(* PLC project Claude2.project, CODESYS CODESYS V3.5 SP20 *)
(* stored: creationDateTime 2026-10-26T14:12:36.8389124, modificationDateTime 2026-10-26T14:11:59.3278775 *)

(* values of E_MachineState: INIT: Inicialização; STOPPED: Parada, sem alarme; HOMING: Referenciamento dos eixos; RUNNING: Ciclo automático; ALARM: Alarme pendente: parada segura; ESTOP: Emergência/porta aberta: sobrepõe tudo *)

{attribute 'qualified_only'}
{attribute 'strict'}
TYPE E_MachineState : (INIT := 0, STOPPED := 10, HOMING := 20, RUNNING := 30, ALARM := 90, ESTOP := 99);
END_TYPE

TYPE ST_Component : STRUCT
  sRef : STRING(20);  (* Designador do componente *)
  rPickX : REAL;  (* Posição de coleta (alimentador) X [mm] *)
  rPickY : REAL;  (* Posição de coleta (alimentador) Y [mm] *)
  rPlaceX : REAL;  (* Posição de montagem X [mm] *)
  rPlaceY : REAL;  (* Posição de montagem Y [mm] *)
  rPlaceTheta : REAL;  (* Ângulo de montagem [graus] *)
END_STRUCT;
END_TYPE

TYPE ST_Recipe : STRUCT
  sName : STRING(30);  (* Nome da receita *)
  iCount : INT;  (* Quantidade de componentes *)
  aComp : ARRAY[1..c_MAX_COMP] OF ST_Component;  (* Lista de componentes *)
END_STRUCT;
END_TYPE

FUNCTION F_InRange : BOOL
  VAR_INPUT
    rValue : REAL;
    rMin : REAL;
    rMax : REAL;
  END_VAR

                  (* Verifica se o valor está dentro da faixa [rMin, rMax] *)
F_InRange := (rValue >= rMin) AND (rValue <= rMax);
                
END_FUNCTION

FUNCTION_BLOCK FB_PneumaticCyl
  VAR_INPUT
    xEnable : BOOL;  (* Habilitação (segurança) *)
    xReset : BOOL;  (* Reset de falha *)
    xCmdExtend : BOOL;  (* TRUE = avançar; FALSE = recuar *)
    xSensExtended : BOOL;
    xSensRetracted : BOOL;
    tMoveTimeout : TIME := TIME#2s0ms;
    tSensorConflict : TIME := TIME#300ms;
  END_VAR
  VAR_OUTPUT
    xValve : BOOL;
    xIsExtended : BOOL;  (* Avançado confirmado: sensor A ligado e B desligado *)
    xIsRetracted : BOOL;  (* Recuado confirmado: sensor B ligado e A desligado *)
    xFault : BOOL;
    iFaultCode : INT;  (* 1 = timeout avanço; 2 = timeout recuo; 3 = sensores em conflito *)
  END_VAR
  VAR
    tonExt : TON;
    tonRet : TON;
    tonBoth : TON;
  END_VAR

                  (* Dupla confirmação *)
xIsExtended  := xSensExtended AND NOT xSensRetracted;
xIsRetracted := xSensRetracted AND NOT xSensExtended;

IF xReset THEN
    xFault := FALSE;
    iFaultCode := 0;
END_IF

(* Supervisão de tempo e de coerência dos sensores *)
tonExt(IN := xEnable AND xValve AND NOT xIsExtended AND NOT xFault, PT := tMoveTimeout);
tonRet(IN := xEnable AND NOT xValve AND NOT xIsRetracted AND NOT xFault, PT := tMoveTimeout);
tonBoth(IN := xEnable AND xSensExtended AND xSensRetracted, PT := tSensorConflict);

IF NOT xFault THEN
    IF tonExt.Q THEN
        xFault := TRUE; iFaultCode := 1;
    ELSIF tonRet.Q THEN
        xFault := TRUE; iFaultCode := 2;
    ELSIF tonBoth.Q THEN
        xFault := TRUE; iFaultCode := 3;
    END_IF
END_IF

(* Saída da válvula: em falha ou sem habilitação, retorna por mola *)
xValve := xEnable AND xCmdExtend AND NOT xFault;
                
END_FUNCTION_BLOCK

FUNCTION_BLOCK FB_VacuumGripper
  VAR_INPUT
    xEnable : BOOL;
    xReset : BOOL;
    xGrip : BOOL;  (* TRUE = segurar; FALSE = liberar *)
    xPressostat : BOOL;
    tConfirm : TIME := TIME#1s0ms;  (* Tempo máximo para confirmar a pega *)
    tDebounce : TIME := TIME#100ms;
    tBlow : TIME := TIME#300ms;
  END_VAR
  VAR_OUTPUT
    xVacValve : BOOL;
    xBlowValve : BOOL;
    xGripOk : BOOL;  (* Pega confirmada *)
    xReleased : BOOL;  (* Liberação confirmada *)
    xPickFail : BOOL;  (* Pega não confirmada no tempo *)
    xGripLoss : BOOL;  (* Perda de vácuo com peça presa *)
  END_VAR
  VAR
    tonOk : TON;
    tonConfirm : TON;
    tonLoss : TON;
    tonRel : TON;
    tonBlow : TON;
    ftGrip : F_TRIG;
    xBlow : BOOL;
    xCarried : BOOL;
  END_VAR

                  xVacValve := xEnable AND xGrip;

(* Janela de sopro após o comando de liberação *)
ftGrip(CLK := xGrip);
IF ftGrip.Q THEN
    xBlow := TRUE;
END_IF
tonBlow(IN := xBlow, PT := tBlow);
IF tonBlow.Q OR xGrip OR NOT xEnable THEN
    xBlow := FALSE;
END_IF
xBlowValve := xBlow AND xEnable;

(* Confirmação da pega *)
tonOk(IN := xGrip AND xPressostat, PT := tDebounce);
xGripOk := tonOk.Q;

(* Falha de pega: vácuo não estabelecido no tempo *)
tonConfirm(IN := xEnable AND xGrip AND NOT xGripOk, PT := tConfirm);
IF tonConfirm.Q THEN
    xPickFail := TRUE;
END_IF
IF xReset OR NOT xGrip THEN
    xPickFail := FALSE;
END_IF

(* Perda de vácuo durante o transporte *)
IF xGripOk THEN
    xCarried := TRUE;
END_IF
IF NOT xGrip THEN
    xCarried := FALSE;
END_IF
tonLoss(IN := xCarried AND xGrip AND NOT xPressostat, PT := tDebounce);
xGripLoss := tonLoss.Q;

(* Confirmação da liberação *)
tonRel(IN := NOT xGrip AND NOT xPressostat, PT := tDebounce);
xReleased := tonRel.Q;
                
END_FUNCTION_BLOCK

FUNCTION_BLOCK FB_AxisCtrl
  VAR_INPUT
    xEnable : BOOL;
    xReset : BOOL;
    xHomeCmd : BOOL;  (* Borda de subida inicia o homing *)
    xMoveCmd : BOOL;  (* Borda de subida inicia o movimento *)
    xHalt : BOOL;  (* Interrompe o movimento em curso *)
    rTarget : REAL;
    rActPos : REAL;
    rSoftMin : REAL;
    rSoftMax : REAL;
    xDriveReady : BOOL;
    xDriveFault : BOOL;
    xDriveHomeDone : BOOL;
    rInPosWindow : REAL := 0.05;
    tSettle : TIME := TIME#100ms;
    tReadyTimeout : TIME := TIME#5s0ms;
    tHomeTimeout : TIME := TIME#1m0s0ms;
    tMoveTimeout : TIME := TIME#15s0ms;
  END_VAR
  VAR_OUTPUT
    xDrivePower : BOOL;
    xDriveHome : BOOL;
    xDriveExecute : BOOL;  (* Pulso de um ciclo *)
    rDriveSetpoint : REAL;
    xHomed : BOOL;
    xInPos : BOOL;
    xBusy : BOOL;
    xAccept : BOOL;  (* Apto a receber comando de homing/movimento *)
    xFault : BOOL;
    iFaultCode : INT;  (* 1 drive não pronto; 2 timeout homing; 3 alvo fora dos limites; 4 timeout movimento; 5 falha do drive; 6 perda de pronto *)
  END_VAR
  VAR
    iState : INT := 0;
    rtHome : R_TRIG;
    rtMove : R_TRIG;
    tonReady : TON;
    tonHome : TON;
    tonMove : TON;
    tonSettle : TON;
    rLastSetpoint : REAL;
    rLatchTarget : REAL;
    xHaltDone : BOOL;
  END_VAR
  VAR CONSTANT
    AS_OFF : INT := 0;
    AS_WAIT_READY : INT := 1;
    AS_UNHOMED : INT := 2;
    AS_HOMING : INT := 3;
    AS_READY : INT := 4;
    AS_START : INT := 5;
    AS_MOVING : INT := 6;
    AS_FAULT : INT := 99;
  END_VAR

                  xDriveExecute := FALSE;
rtHome(CLK := xHomeCmd);
rtMove(CLK := xMoveCmd);

tonReady(IN := (iState = AS_WAIT_READY), PT := tReadyTimeout);
tonHome(IN := (iState = AS_HOMING), PT := tHomeTimeout);
tonMove(IN := (iState = AS_MOVING), PT := tMoveTimeout);
tonSettle(IN := (iState = AS_MOVING) AND (ABS(rActPos - rLastSetpoint) <= rInPosWindow),
          PT := tSettle);

(* Supervisão geral *)
IF iState <> AS_FAULT THEN
    IF NOT xEnable THEN
        iState := AS_OFF;
    ELSIF iState >= AS_WAIT_READY THEN
        IF xDriveFault THEN
            iFaultCode := 5; iState := AS_FAULT;
        ELSIF (iState >= AS_UNHOMED) AND NOT xDriveReady THEN
            iFaultCode := 6; iState := AS_FAULT;
        END_IF
    END_IF
END_IF

CASE iState OF
    AS_OFF:
        xHomed := FALSE;
        IF xEnable THEN
            iState := AS_WAIT_READY;
        END_IF

    AS_WAIT_READY:
        IF xDriveReady THEN
            iState := AS_UNHOMED;
        ELSIF tonReady.Q THEN
            iFaultCode := 1; iState := AS_FAULT;
        END_IF

    AS_UNHOMED:
        IF rtHome.Q THEN
            iState := AS_HOMING;
        END_IF

    AS_HOMING:
        IF xDriveHomeDone THEN
            xHomed := TRUE;
            rLastSetpoint := rActPos;
            iState := AS_READY;
        ELSIF tonHome.Q THEN
            iFaultCode := 2; iState := AS_FAULT;
        END_IF

    AS_READY:
        IF rtHome.Q THEN
            xHomed := FALSE;
            iState := AS_HOMING;
        ELSIF rtMove.Q THEN
            IF (rTarget < rSoftMin) OR (rTarget > rSoftMax) THEN
                iFaultCode := 3; iState := AS_FAULT;
            ELSE
                rLatchTarget := rTarget;
                iState := AS_START;
            END_IF
        END_IF

    AS_START:
        rDriveSetpoint := rLatchTarget;
        rLastSetpoint := rLatchTarget;
        xDriveExecute := TRUE;
        iState := AS_MOVING;

    AS_MOVING:
        IF xHalt AND NOT xHaltDone THEN
            (* Parada: novo alvo = posição atual *)
            rDriveSetpoint := rActPos;
            rLastSetpoint := rActPos;
            xDriveExecute := TRUE;
            xHaltDone := TRUE;
        END_IF
        IF tonSettle.Q THEN
            iState := AS_READY;
        ELSIF tonMove.Q THEN
            iFaultCode := 4; iState := AS_FAULT;
        END_IF

    AS_FAULT:
        xHomed := FALSE;
        IF xReset AND NOT xDriveFault THEN
            iFaultCode := 0;
            iState := AS_OFF;
        END_IF
END_CASE

IF iState <> AS_MOVING THEN
    xHaltDone := FALSE;
END_IF

(* Saídas *)
xDrivePower := (iState >= AS_WAIT_READY) AND (iState <> AS_FAULT);
xDriveHome  := (iState = AS_HOMING);
xBusy       := (iState = AS_HOMING) OR (iState = AS_START) OR (iState = AS_MOVING);
xAccept     := (iState = AS_UNHOMED) OR (iState = AS_READY);
xInPos      := (iState = AS_READY) AND xHomed AND (ABS(rActPos - rLastSetpoint) <= rInPosWindow);
xFault      := (iState = AS_FAULT);
                
END_FUNCTION_BLOCK

FUNCTION_BLOCK FB_Conveyor
  VAR_INPUT
    xEnable : BOOL;  (* Ciclo automático liberado *)
    xReset : BOOL;
    xClearZones : BOOL;  (* Ressincroniza zonas pelos sensores *)
    xSensZ1 : BOOL;
    xSensZ2 : BOOL;
    xSensZ3 : BOOL;
    xUpBoardAvail : BOOL;  (* SMEMA a montante: placa disponível *)
    xDownMachineReady : BOOL;  (* SMEMA a jusante: máquina pronta *)
    xAsmDone : BOOL;  (* Montagem concluída: libera a zona 2 *)
    xInspDone : BOOL;  (* Inspeção concluída: libera a zona 3 *)
    tTransferTimeout : TIME := TIME#15s0ms;
    tSensorFilter : TIME := TIME#50ms;
    tClearDelay : TIME := TIME#500ms;
  END_VAR
  VAR_OUTPUT
    xMotor1 : BOOL;
    xMotor2 : BOOL;
    xMotor3 : BOOL;
    xUpMachineReady : BOOL;  (* SMEMA a montante: máquina pronta *)
    xDownBoardAvail : BOOL;  (* SMEMA a jusante: placa disponível *)
    xBoardInAsm : BOOL;
    xBoardInInsp : BOOL;
    xFault : BOOL;
  END_VAR
  VAR
    iZ1 : INT;  (* Estado de cada zona *)
    iZ2 : INT;  (* Estado de cada zona *)
    iZ3 : INT;  (* Estado de cada zona *)
    tonP1 : TON;  (* Presença filtrada *)
    tonP2 : TON;  (* Presença filtrada *)
    tonP3 : TON;  (* Presença filtrada *)
    tonA1 : TON;  (* Ausência filtrada *)
    tonA2 : TON;  (* Ausência filtrada *)
    tonA3 : TON;  (* Ausência filtrada *)
    tonT1 : TON;  (* Timeout de movimento *)
    tonT2 : TON;  (* Timeout de movimento *)
    tonT3 : TON;  (* Timeout de movimento *)
    xP1 : BOOL;
    xP2 : BOOL;
    xP3 : BOOL;
    xA1 : BOOL;
    xA2 : BOOL;
    xA3 : BOOL;
    xActive : BOOL;
  END_VAR
  VAR CONSTANT
    ZS_EMPTY : INT := 0;
    ZS_RECV : INT := 1;  (* Recebendo placa *)
    ZS_OCC : INT := 2;  (* Placa posicionada *)
    ZS_SEND : INT := 3;  (* Enviando placa *)
  END_VAR

                  (* Filtros dos sensores *)
tonP1(IN := xSensZ1, PT := tSensorFilter);   xP1 := tonP1.Q;
tonP2(IN := xSensZ2, PT := tSensorFilter);   xP2 := tonP2.Q;
tonP3(IN := xSensZ3, PT := tSensorFilter);   xP3 := tonP3.Q;
tonA1(IN := NOT xSensZ1, PT := tClearDelay); xA1 := tonA1.Q;
tonA2(IN := NOT xSensZ2, PT := tClearDelay); xA2 := tonA2.Q;
tonA3(IN := NOT xSensZ3, PT := tClearDelay); xA3 := tonA3.Q;

IF xReset THEN
    xFault := FALSE;
END_IF

(* Ressincronização: considera placa posicionada onde houver sensor ativo *)
IF xClearZones THEN
    IF xSensZ1 THEN iZ1 := ZS_OCC; ELSE iZ1 := ZS_EMPTY; END_IF
    IF xSensZ2 THEN iZ2 := ZS_OCC; ELSE iZ2 := ZS_EMPTY; END_IF
    IF xSensZ3 THEN iZ3 := ZS_OCC; ELSE iZ3 := ZS_EMPTY; END_IF
    xFault := FALSE;
END_IF

(* Timeout de transferência (motores acionados no ciclo anterior) *)
tonT1(IN := xMotor1, PT := tTransferTimeout);
tonT2(IN := xMotor2, PT := tTransferTimeout);
tonT3(IN := xMotor3, PT := tTransferTimeout);
IF tonT1.Q OR tonT2.Q OR tonT3.Q THEN
    xFault := TRUE;
END_IF

xActive := xEnable AND NOT xFault;

(* ---------- Zona 1: entrada ---------- *)
CASE iZ1 OF
    ZS_EMPTY:
        IF xActive AND xUpBoardAvail THEN
            iZ1 := ZS_RECV;
        END_IF
    ZS_RECV:
        IF xP1 THEN
            iZ1 := ZS_OCC;
        END_IF
    ZS_OCC:
        IF xActive AND (iZ2 = ZS_EMPTY) THEN
            iZ1 := ZS_SEND;
            iZ2 := ZS_RECV;     (* Transferência 1 -> 2 *)
        END_IF
    ZS_SEND:
        IF (iZ2 = ZS_OCC) AND xA1 THEN
            iZ1 := ZS_EMPTY;
        END_IF
END_CASE

(* ---------- Zona 2: montagem ---------- *)
CASE iZ2 OF
    ZS_EMPTY:
        ;
    ZS_RECV:
        IF xP2 THEN
            iZ2 := ZS_OCC;
        END_IF
    ZS_OCC:
        IF xActive AND xAsmDone AND (iZ3 = ZS_EMPTY) THEN
            iZ2 := ZS_SEND;
            iZ3 := ZS_RECV;     (* Transferência 2 -> 3 *)
        END_IF
    ZS_SEND:
        IF (iZ3 = ZS_OCC) AND xA2 THEN
            iZ2 := ZS_EMPTY;
        END_IF
END_CASE

(* ---------- Zona 3: saída / inspeção ---------- *)
CASE iZ3 OF
    ZS_EMPTY:
        ;
    ZS_RECV:
        IF xP3 THEN
            iZ3 := ZS_OCC;
        END_IF
    ZS_OCC:
        IF xActive AND xInspDone THEN
            iZ3 := ZS_SEND;
        END_IF
    ZS_SEND:
        IF xA3 THEN
            iZ3 := ZS_EMPTY;
        END_IF
END_CASE

(* ---------- Saídas (calculadas após a lógica de estados) ---------- *)
xMotor1 := xActive AND ((iZ1 = ZS_RECV) OR (iZ1 = ZS_SEND));
xMotor2 := xActive AND ((iZ2 = ZS_RECV) OR (iZ2 = ZS_SEND));
xMotor3 := xActive AND ((iZ3 = ZS_RECV) OR ((iZ3 = ZS_SEND) AND xDownMachineReady));

xUpMachineReady := xActive AND ((iZ1 = ZS_EMPTY) OR (iZ1 = ZS_RECV));
xDownBoardAvail := (iZ3 = ZS_SEND);
xBoardInAsm     := (iZ2 = ZS_OCC);
xBoardInInsp    := (iZ3 = ZS_OCC);
                
END_FUNCTION_BLOCK

FUNCTION_BLOCK FB_HmiWatchdog
  VAR_INPUT
    iHeartbeat : UINT;
    tTimeout : TIME := TIME#3s0ms;
  END_VAR
  VAR_OUTPUT
    xOk : BOOL;
    xLost : BOOL;
  END_VAR
  VAR
    uiLast : UINT;
    xFirst : BOOL := TRUE;
    xChanged : BOOL;
    tonLoss : TON;
  END_VAR

                  IF xFirst THEN
    uiLast := iHeartbeat;
    xFirst := FALSE;
END_IF

xChanged := (iHeartbeat <> uiLast);
uiLast := iHeartbeat;

tonLoss(IN := NOT xChanged, PT := tTimeout);
xLost := tonLoss.Q;
xOk := NOT tonLoss.Q;
                
END_FUNCTION_BLOCK

FUNCTION_BLOCK FB_Alarm
  VAR_INPUT
    xCondition : BOOL;  (* Condição de alarme (nível ou pulso) *)
    xAck : BOOL;
    xReset : BOOL;
  END_VAR
  VAR_OUTPUT
    xActive : BOOL;  (* Alarme retido *)
    xAcked : BOOL;
  END_VAR
  VAR
    rtCond : R_TRIG;
    rtAck : R_TRIG;
    rtRst : R_TRIG;
  END_VAR

                  rtCond(CLK := xCondition);
rtAck(CLK := xAck);
rtRst(CLK := xReset);

IF rtCond.Q THEN
    xActive := TRUE;
    xAcked := FALSE;
END_IF

IF rtAck.Q AND xActive THEN
    xAcked := TRUE;
END_IF

(* Reset só é aceito com alarme reconhecido e condição normalizada *)
IF rtRst.Q AND xActive AND xAcked AND NOT xCondition THEN
    xActive := FALSE;
    xAcked := FALSE;
END_IF
                
END_FUNCTION_BLOCK

FUNCTION_BLOCK FB_Recipe
  VAR_INPUT
    xRequest : BOOL;  (* Borda de subida solicita a troca *)
    iRequested : INT;
    xMachineStopped : BOOL;
    rXMin : REAL;
    rXMax : REAL;
    rYMin : REAL;
    rYMax : REAL;
  END_VAR
  VAR_IN_OUT
    aRecipes : ARRAY[1..c_NUM_RECIPES] OF ST_Recipe;
  END_VAR
  VAR_OUTPUT
    iActive : INT;
    xValid : BOOL;
    xRejected : BOOL;
  END_VAR
  VAR
    rtReq : R_TRIG;
    i : INT;
    xOk : BOOL;
    stC : ST_Component;
  END_VAR

                  rtReq(CLK := xRequest);

IF rtReq.Q THEN
    IF xMachineStopped AND (iRequested >= 1) AND (iRequested <= c_NUM_RECIPES) THEN
        iActive := iRequested;
        xRejected := FALSE;
    ELSE
        xRejected := TRUE;
    END_IF
END_IF
IF NOT xRequest THEN
    xRejected := FALSE;
END_IF

(* Validação da receita ativa *)
xOk := (iActive >= 1) AND (iActive <= c_NUM_RECIPES);
IF xOk THEN
    xOk := (aRecipes[iActive].iCount >= 1) AND (aRecipes[iActive].iCount <= c_MAX_COMP);
END_IF
IF xOk THEN
    FOR i := 1 TO aRecipes[iActive].iCount DO
        stC := aRecipes[iActive].aComp[i];
        IF NOT (F_InRange(stC.rPickX, rXMin, rXMax)
            AND F_InRange(stC.rPickY, rYMin, rYMax)
            AND F_InRange(stC.rPlaceX, rXMin, rXMax)
            AND F_InRange(stC.rPlaceY, rYMin, rYMax)
            AND F_InRange(stC.rPlaceTheta, -180.0, 180.0)) THEN
            xOk := FALSE;
            EXIT;
        END_IF
    END_FOR
END_IF
xValid := xOk;
                
END_FUNCTION_BLOCK

PROGRAM PRG_Safety
  VAR
    tonRearm : TON;
    fbHmi : FB_HmiWatchdog;
  END_VAR

                  (* Perda imediata; rearme somente após 500 ms de condição normal *)
tonRearm(IN := xEStopOk AND xDoorClosed, PT := T#500MS);
xSafetyOk := tonRearm.Q;

(* Heartbeat da IHM *)
fbHmi(iHeartbeat := iHmiHeartbeat, tTimeout := tHmiTimeout);
xHmiOk := fbHmi.xOk;
                
END_PROGRAM

PROGRAM PRG_Alarms
  VAR
    fbAlarm : ARRAY[1..15] OF FB_Alarm;
    aCond : ARRAY[1..15] OF BOOL;
    i : INT;
  END_VAR

                  (* Condições de alarme *)
aCond[c_ALM_ESTOP]       := NOT xEStopOk;
aCond[c_ALM_DOOR]        := NOT xDoorClosed;
aCond[c_ALM_HMI]         := NOT xHmiOk;
aCond[c_ALM_CONVEYOR]    := xConveyorFault;
FOR i := 1 TO 4 DO
    aCond[c_ALM_AXIS_X + i - 1] := xAxisFault[i];
END_FOR
aCond[c_ALM_CLAMP]       := xClampFault;
aCond[c_ALM_STOPPER]     := xStopperFault;
aCond[c_ALM_PICK_FAIL]   := xPickFail;
aCond[c_ALM_VAC_LOSS]    := xGripLoss;
aCond[c_ALM_AOI_TIMEOUT] := xAoiTimeout;
aCond[c_ALM_RECIPE]      := xStartRefusedRecipe;
aCond[c_ALM_Z_INTERLOCK] := xZInterlockFault;

(* Processamento e consolidação *)
xAnyAlarm := FALSE;
xAnyUnacked := FALSE;
FOR i := 1 TO c_NUM_ALARMS DO
    fbAlarm[i](xCondition := aCond[i], xAck := xCmdAck, xReset := xCmdReset);
    xAlarmActive[i] := fbAlarm[i].xActive;
    xAlarmAcked[i]  := fbAlarm[i].xAcked;
    IF fbAlarm[i].xActive THEN
        xAnyAlarm := TRUE;
        IF NOT fbAlarm[i].xAcked THEN
            xAnyUnacked := TRUE;
        END_IF
    END_IF
END_FOR
                
END_PROGRAM

PROGRAM PRG_Main
  VAR
    fbRecipe : FB_Recipe;
    rtReset : R_TRIG;
    rtStart : R_TRIG;
    rtStop : R_TRIG;
    rtHome : R_TRIG;
    xStopped : BOOL;
  END_VAR

                  rtReset(CLK := xCmdReset);
rtStart(CLK := xCmdStart);
rtStop(CLK := xCmdStop);
rtHome(CLK := xCmdHome);
xResetPulse := rtReset.Q;
xStartRefusedRecipe := FALSE;

(* Receitas: troca somente com a máquina parada *)
xStopped := (eMachineState <> E_MachineState.RUNNING) AND (eMachineState <> E_MachineState.HOMING);
fbRecipe(xRequest := xCmdRecipeSel,
         iRequested := iRecipeReq,
         xMachineStopped := xStopped,
         rXMin := rAxisMin[c_AX_X], rXMax := rAxisMax[c_AX_X],
         rYMin := rAxisMin[c_AX_Y], rYMax := rAxisMax[c_AX_Y],
         aRecipes := aRecipes);
iRecipeActive   := fbRecipe.iActive;
xRecipeValid    := fbRecipe.xValid;
xRecipeRejected := fbRecipe.xRejected;

(* Emergência e porta sobrepõem qualquer estado *)
IF NOT xSafetyOk THEN
    eMachineState := E_MachineState.ESTOP;
ELSE
    CASE eMachineState OF
        E_MachineState.INIT, E_MachineState.ESTOP:
            IF xAnyAlarm THEN
                eMachineState := E_MachineState.ALARM;
            ELSE
                eMachineState := E_MachineState.STOPPED;
            END_IF

        E_MachineState.STOPPED:
            IF xAnyAlarm THEN
                eMachineState := E_MachineState.ALARM;
            ELSIF rtHome.Q THEN
                eMachineState := E_MachineState.HOMING;
            ELSIF rtStart.Q THEN
                IF NOT xAllHomed THEN
                    ;   (* Partida ignorada: eixos não referenciados *)
                ELSIF NOT xRecipeValid THEN
                    xStartRefusedRecipe := TRUE;
                ELSE
                    eMachineState := E_MachineState.RUNNING;
                END_IF
            END_IF

        E_MachineState.HOMING:
            IF xAnyAlarm THEN
                eMachineState := E_MachineState.ALARM;
            ELSIF xHomeSeqDone THEN
                eMachineState := E_MachineState.STOPPED;
            END_IF

        E_MachineState.RUNNING:
            IF xAnyAlarm THEN
                eMachineState := E_MachineState.ALARM;
            ELSIF rtStop.Q THEN
                eMachineState := E_MachineState.STOPPED;
            END_IF

        E_MachineState.ALARM:
            IF NOT xAnyAlarm THEN
                eMachineState := E_MachineState.STOPPED;
            END_IF
    END_CASE
END_IF

(* Habilitações derivadas do estado *)
xDrivesEnable := xSafetyOk;
xAutoEnable   := (eMachineState = E_MachineState.RUNNING);
xMotionRun    := xAutoEnable OR (eMachineState = E_MachineState.HOMING);
xHomeReq      := (eMachineState = E_MachineState.HOMING);
                
END_PROGRAM

PROGRAM PRG_Motion
  VAR
    fbAx : ARRAY[1..4] OF FB_AxisCtrl;
    xCmdHomeAx : ARRAY[1..4] OF BOOL;
    xCmdMoveAx : ARRAY[1..4] OF BOOL;
    rTgt : ARRAY[1..4] OF REAL;
    iSvc : INT := 0;
    i : INT;
    xZSafe : BOOL;
    xAccXYT : BOOL;
    xInPosXYT : BOOL;
    xHomedXYT : BOOL;
  END_VAR
  VAR CONSTANT
    SV_IDLE : INT := 0;
    SV_HOME_Z : INT := 10;
    SV_HOME_Z_W : INT := 11;
    SV_Z_SAFE : INT := 12;
    SV_Z_SAFE_W : INT := 13;
    SV_HOME_XYT : INT := 14;
    SV_HOME_XYT_W : INT := 15;
    SV_PARK : INT := 16;
    SV_PARK_W : INT := 17;
    SV_XYT_GO : INT := 20;
    SV_XYT_W : INT := 21;
    SV_Z_GO : INT := 30;
    SV_Z_W : INT := 31;
  END_VAR

                  (* Comandos são pulsos de um ciclo *)
FOR i := 1 TO 4 DO
    xCmdHomeAx[i] := FALSE;
    xCmdMoveAx[i] := FALSE;
END_FOR
xZInterlockFault := FALSE;

xZSafe    := rAxisActPos[c_AX_Z] >= (rZSafe - rZTol);
xAccXYT   := fbAx[c_AX_X].xAccept AND fbAx[c_AX_Y].xAccept AND fbAx[c_AX_T].xAccept;
xInPosXYT := fbAx[c_AX_X].xInPos  AND fbAx[c_AX_Y].xInPos  AND fbAx[c_AX_T].xInPos;
xHomedXYT := fbAx[c_AX_X].xHomed  AND fbAx[c_AX_Y].xHomed  AND fbAx[c_AX_T].xHomed;

IF (NOT xMotionRun) OR xMotionFault THEN
    (* Aborta os serviços *)
    iSvc := SV_IDLE;
    xXYTDone := FALSE;
    xZDone := FALSE;
    xHomeSeqDone := FALSE;
ELSE
    CASE iSvc OF
        SV_IDLE:
            xXYTDone     := xXYTDone AND xMoveXYTReq;
            xZDone       := xZDone AND xMoveZReq;
            xHomeSeqDone := xHomeSeqDone AND xHomeReq;
            IF xHomeReq AND NOT xHomeSeqDone THEN
                iSvc := SV_HOME_Z;
            ELSIF xMoveXYTReq AND NOT xXYTDone AND xAllHomed THEN
                IF xZSafe THEN
                    iSvc := SV_XYT_GO;
                ELSE
                    xZInterlockFault := TRUE;   (* XYθ só com Z na altura segura *)
                END_IF
            ELSIF xMoveZReq AND NOT xZDone AND xAllHomed THEN
                iSvc := SV_Z_GO;
            END_IF

        (* ----- Sequência de homing ----- *)
        SV_HOME_Z:
            IF fbAx[c_AX_Z].xAccept THEN
                xCmdHomeAx[c_AX_Z] := TRUE;
                iSvc := SV_HOME_Z_W;
            END_IF
        SV_HOME_Z_W:
            IF fbAx[c_AX_Z].xHomed AND fbAx[c_AX_Z].xInPos THEN
                iSvc := SV_Z_SAFE;
            END_IF
        SV_Z_SAFE:
            rTgt[c_AX_Z] := rZSafe;
            IF fbAx[c_AX_Z].xAccept THEN
                xCmdMoveAx[c_AX_Z] := TRUE;
                iSvc := SV_Z_SAFE_W;
            END_IF
        SV_Z_SAFE_W:
            IF fbAx[c_AX_Z].xInPos THEN
                iSvc := SV_HOME_XYT;
            END_IF
        SV_HOME_XYT:
            IF xAccXYT THEN
                xCmdHomeAx[c_AX_X] := TRUE;
                xCmdHomeAx[c_AX_Y] := TRUE;
                xCmdHomeAx[c_AX_T] := TRUE;
                iSvc := SV_HOME_XYT_W;
            END_IF
        SV_HOME_XYT_W:
            IF xHomedXYT AND xInPosXYT THEN
                iSvc := SV_PARK;
            END_IF
        SV_PARK:
            rTgt[c_AX_X] := rParkX;
            rTgt[c_AX_Y] := rParkY;
            rTgt[c_AX_T] := rParkT;
            IF xAccXYT THEN
                xCmdMoveAx[c_AX_X] := TRUE;
                xCmdMoveAx[c_AX_Y] := TRUE;
                xCmdMoveAx[c_AX_T] := TRUE;
                iSvc := SV_PARK_W;
            END_IF
        SV_PARK_W:
            IF xInPosXYT THEN
                xHomeSeqDone := TRUE;
                iSvc := SV_IDLE;
            END_IF

        (* ----- Movimento XYθ ----- *)
        SV_XYT_GO:
            rTgt[c_AX_X] := rTgtX;
            rTgt[c_AX_Y] := rTgtY;
            rTgt[c_AX_T] := rTgtT;
            IF xAccXYT THEN
                xCmdMoveAx[c_AX_X] := TRUE;
                xCmdMoveAx[c_AX_Y] := TRUE;
                xCmdMoveAx[c_AX_T] := TRUE;
                iSvc := SV_XYT_W;
            END_IF
        SV_XYT_W:
            IF xInPosXYT THEN
                xXYTDone := TRUE;
                iSvc := SV_IDLE;
            END_IF

        (* ----- Movimento Z ----- *)
        SV_Z_GO:
            rTgt[c_AX_Z] := rTgtZ;
            IF fbAx[c_AX_Z].xAccept THEN
                xCmdMoveAx[c_AX_Z] := TRUE;
                iSvc := SV_Z_W;
            END_IF
        SV_Z_W:
            IF fbAx[c_AX_Z].xInPos THEN
                xZDone := TRUE;
                iSvc := SV_IDLE;
            END_IF
    END_CASE
END_IF

(* Execução dos eixos *)
xAllHomed := TRUE;
xMotionFault := FALSE;
FOR i := 1 TO 4 DO
    fbAx[i](xEnable        := xDrivesEnable,
            xReset         := xResetPulse,
            xHomeCmd       := xCmdHomeAx[i],
            xMoveCmd       := xCmdMoveAx[i],
            xHalt          := (NOT xMotionRun) OR xMotionFault,
            rTarget        := rTgt[i],
            rActPos        := rAxisActPos[i],
            rSoftMin       := rAxisMin[i],
            rSoftMax       := rAxisMax[i],
            xDriveReady    := xAxisDriveReady[i],
            xDriveFault    := xAxisDriveFault[i],
            xDriveHomeDone := xAxisHomeDone[i]);

    xAxisPower[i]    := fbAx[i].xDrivePower;
    xAxisHome[i]     := fbAx[i].xDriveHome;
    xAxisExecute[i]  := fbAx[i].xDriveExecute;
    rAxisSetpoint[i] := fbAx[i].rDriveSetpoint;
    xAxisFault[i]    := fbAx[i].xFault;

    xAllHomed := xAllHomed AND fbAx[i].xHomed;
    IF fbAx[i].xFault THEN
        xMotionFault := TRUE;
    END_IF
END_FOR
                
END_PROGRAM

PROGRAM PRG_Conveyor
  VAR
    fbConv : FB_Conveyor;
  END_VAR

                  fbConv(xEnable           := xAutoEnable AND xSafetyOk,
       xReset            := xResetPulse,
       xClearZones       := xCmdClearZones AND NOT xAutoEnable,
       xSensZ1           := xSensZ1,
       xSensZ2           := xSensZ2,
       xSensZ3           := xSensZ3,
       xUpBoardAvail     := xSmemaUpAvail,
       xDownMachineReady := xSmemaDownReady,
       xAsmDone          := xAsmDone,
       xInspDone         := xInspDone,
       tTransferTimeout  := tConvTimeout);

xMotor1         := fbConv.xMotor1;
xMotor2         := fbConv.xMotor2;
xMotor3         := fbConv.xMotor3;
xSmemaUpReady   := fbConv.xUpMachineReady;
xSmemaDownAvail := fbConv.xDownBoardAvail;
xBoardInAsm     := fbConv.xBoardInAsm;
xBoardInInsp    := fbConv.xBoardInInsp;
xConveyorFault  := fbConv.xFault;
                
END_PROGRAM

PROGRAM PRG_PickPlace
  VAR
    iStep : INT := 0;
    iComp : INT := 1;
    iCount : INT;
    stCur : ST_Component;
    xGripCmd : BOOL;
    xClampCmd : BOOL;
    fbClamp : FB_PneumaticCyl;
    fbVac : FB_VacuumGripper;
    rtBoard : R_TRIG;
  END_VAR
  VAR CONSTANT
    S_IDLE : INT := 0;
    S_CLAMP : INT := 10;
    S_LIFT : INT := 15;
    S_PICK_XY : INT := 20;
    S_PICK_DOWN : INT := 30;
    S_GRIP : INT := 40;
    S_PICK_UP : INT := 50;
    S_PLACE_XY : INT := 60;
    S_PLACE_DOWN : INT := 70;
    S_RELEASE : INT := 80;
    S_PLACE_UP : INT := 90;
    S_NEXT : INT := 100;
    S_UNCLAMP : INT := 110;
    S_DONE : INT := 120;
  END_VAR

                  (* Nova placa na zona de montagem: reinicia a lista de componentes *)
rtBoard(CLK := xBoardInAsm);
IF rtBoard.Q THEN
    iComp := 1;
END_IF

(* Componente corrente da receita ativa *)
IF xRecipeValid AND (iRecipeActive >= 1) AND (iRecipeActive <= c_NUM_RECIPES) THEN
    iCount := aRecipes[iRecipeActive].iCount;
    IF (iComp >= 1) AND (iComp <= iCount) THEN
        stCur := aRecipes[iRecipeActive].aComp[iComp];
    END_IF
ELSE
    iCount := 0;
END_IF

IF NOT xAutoEnable THEN
    (* Aborto seguro: cancela requisições, libera vácuo e grampo *)
    xMoveXYTReq := FALSE;
    xMoveZReq   := FALSE;
    xGripCmd    := FALSE;
    xClampCmd   := FALSE;
    iStep       := S_IDLE;
ELSE
    CASE iStep OF
        S_IDLE:
            IF xAsmDone THEN
                IF NOT xBoardInAsm THEN
                    xAsmDone := FALSE;
                END_IF
            ELSIF xBoardInAsm AND (iCount > 0) THEN
                IF iComp > iCount THEN
                    iStep := S_UNCLAMP;     (* Todos colocados antes do aborto *)
                ELSE
                    iStep := S_CLAMP;
                END_IF
            END_IF

        S_CLAMP:
            xClampCmd := TRUE;
            IF fbClamp.xIsExtended THEN
                iStep := S_LIFT;
            END_IF

        S_LIFT:     (* Garante Z seguro antes de qualquer movimento XY *)
            rTgtZ := rZSafe;
            xMoveZReq := TRUE;
            IF xZDone THEN
                xMoveZReq := FALSE;
                iStep := S_PICK_XY;
            END_IF

        S_PICK_XY:
            rTgtX := stCur.rPickX;
            rTgtY := stCur.rPickY;
            rTgtT := 0.0;
            xMoveXYTReq := TRUE;
            IF xXYTDone THEN
                xMoveXYTReq := FALSE;
                iStep := S_PICK_DOWN;
            END_IF

        S_PICK_DOWN:
            rTgtZ := rZPick;
            xMoveZReq := TRUE;
            IF xZDone THEN
                xMoveZReq := FALSE;
                iStep := S_GRIP;
            END_IF

        S_GRIP:     (* Confirma a pega pelo pressostato *)
            xGripCmd := TRUE;
            IF fbVac.xGripOk THEN
                iStep := S_PICK_UP;
            END_IF

        S_PICK_UP:
            rTgtZ := rZSafe;
            xMoveZReq := TRUE;
            IF xZDone THEN
                xMoveZReq := FALSE;
                iStep := S_PLACE_XY;
            END_IF

        S_PLACE_XY:
            rTgtX := stCur.rPlaceX;
            rTgtY := stCur.rPlaceY;
            rTgtT := stCur.rPlaceTheta;
            xMoveXYTReq := TRUE;
            IF xXYTDone THEN
                xMoveXYTReq := FALSE;
                iStep := S_PLACE_DOWN;
            END_IF

        S_PLACE_DOWN:
            rTgtZ := rZPlace;
            xMoveZReq := TRUE;
            IF xZDone THEN
                xMoveZReq := FALSE;
                iStep := S_RELEASE;
            END_IF

        S_RELEASE:
            xGripCmd := FALSE;
            IF fbVac.xReleased THEN
                iStep := S_PLACE_UP;
            END_IF

        S_PLACE_UP:
            rTgtZ := rZSafe;
            xMoveZReq := TRUE;
            IF xZDone THEN
                xMoveZReq := FALSE;
                iStep := S_NEXT;
            END_IF

        S_NEXT:
            iComp := iComp + 1;
            IF iComp > iCount THEN
                iStep := S_UNCLAMP;
            ELSE
                iStep := S_PICK_XY;
            END_IF

        S_UNCLAMP:
            xClampCmd := FALSE;
            IF fbClamp.xIsRetracted THEN
                iStep := S_DONE;
            END_IF

        S_DONE:     (* Libera a placa para a esteira *)
            xAsmDone := TRUE;
            IF NOT xBoardInAsm THEN
                xAsmDone := FALSE;
                iStep := S_IDLE;
            END_IF
    END_CASE
END_IF

(* Atuadores *)
fbClamp(xEnable         := xSafetyOk,
        xReset          := xResetPulse,
        xCmdExtend      := xClampCmd,
        xSensExtended   := xClampExtended,
        xSensRetracted  := xClampRetracted,
        tMoveTimeout    := tCylTimeout);
xClampValve := fbClamp.xValve;
xClampFault := fbClamp.xFault;

fbVac(xEnable     := xSafetyOk,
      xReset      := xResetPulse,
      xGrip       := xGripCmd,
      xPressostat := xVacuumOk,
      tConfirm    := tVacConfirm);
xVacValve  := fbVac.xVacValve;
xBlowValve := fbVac.xBlowValve;
xPickFail  := fbVac.xPickFail;
xGripLoss  := fbVac.xGripLoss;
                
END_PROGRAM

PROGRAM PRG_AOI
  VAR
    iStep : INT := 0;
    iFails : INT;
    xPass : BOOL;
    xReject : BOOL;
    xStopExtend : BOOL;
    fbStop : FB_PneumaticCyl;
    tonRes : TON;
    tonRel : TON;
    rtResetCnt : R_TRIG;
  END_VAR
  VAR CONSTANT
    A_IDLE : INT := 0;
    A_WAIT_STOP : INT := 10;
    A_WAIT_RESULT : INT := 20;
    A_WAIT_RELEASE : INT := 30;
    A_RETRACT : INT := 40;
    A_DONE : INT := 50;
  END_VAR

                  (* Zerar contadores somente com o ciclo automático parado *)
rtResetCnt(CLK := xCmdResetCounters);
IF rtResetCnt.Q AND NOT xAutoEnable THEN
    diBoardsProduced := 0;
    diBoardsRejected := 0;
END_IF

(* Supervisão de tempo da AOI *)
tonRes(IN := (iStep = A_WAIT_RESULT), PT := tAoiTimeout);
tonRel(IN := (iStep = A_WAIT_RELEASE), PT := tAoiTimeout);
xAoiTimeout := tonRes.Q OR tonRel.Q;

IF NOT xAutoEnable THEN
    xAoiTrigger := FALSE;
    iStep := A_IDLE;
ELSE
    CASE iStep OF
        A_IDLE:
            IF xInspDone THEN
                IF NOT xBoardInInsp THEN
                    xInspDone := FALSE;
                END_IF
            ELSIF xBoardInInsp THEN
                iFails := 0;
                iStep := A_WAIT_STOP;
            END_IF

        A_WAIT_STOP:    (* Placa contra o batente avançado *)
            IF fbStop.xIsExtended THEN
                iStep := A_WAIT_RESULT;
            END_IF

        A_WAIT_RESULT:
            xAoiTrigger := TRUE;
            IF xAoiDone THEN
                xPass := xAoiPass;
                xAoiTrigger := FALSE;
                iStep := A_WAIT_RELEASE;
            END_IF

        A_WAIT_RELEASE: (* Aguarda a AOI baixar o resultado antes de decidir *)
            IF NOT xAoiDone THEN
                IF xPass THEN
                    xReject := FALSE;
                    iStep := A_RETRACT;
                ELSE
                    iFails := iFails + 1;
                    IF iFails > c_AOI_MAX_RETRY THEN
                        xReject := TRUE;
                        iStep := A_RETRACT;
                    ELSE
                        iStep := A_WAIT_RESULT;     (* Nova tentativa *)
                    END_IF
                END_IF
            END_IF

        A_RETRACT:      (* Recua o batente e então libera a placa *)
            IF fbStop.xIsRetracted THEN
                diBoardsProduced := diBoardsProduced + 1;
                IF xReject THEN
                    diBoardsRejected := diBoardsRejected + 1;
                END_IF
                xCurBoardRejected := xReject;
                xInspDone := TRUE;
                iStep := A_DONE;
            END_IF

        A_DONE:
            IF NOT xBoardInInsp THEN
                xInspDone := FALSE;
                iStep := A_IDLE;
            END_IF
    END_CASE
END_IF

(* Marca de rejeição acompanha a placa até sair da zona de saída *)
IF NOT xBoardInInsp AND NOT xSmemaDownAvail THEN
    xCurBoardRejected := FALSE;
END_IF
xBoardRejectedOut := xCurBoardRejected;

(* Batente: avançado, exceto durante a liberação da placa *)
xStopExtend := NOT ((iStep = A_RETRACT) OR xInspDone);
fbStop(xEnable        := xSafetyOk,
       xReset         := xResetPulse,
       xCmdExtend     := xStopExtend,
       xSensExtended  := xStopExtended,
       xSensRetracted := xStopRetracted,
       tMoveTimeout   := tCylTimeout);
xStopValve    := fbStop.xValve;
xStopperFault := fbStop.xFault;
                
END_PROGRAM

CONFIGURATION Application
  RESOURCE Application ON PLC
    VAR_GLOBAL CONSTANT  (* GVL_Main - ===================== CONSTANTES ===================== *)
      c_NUM_RECIPES : INT := 3;
      c_MAX_COMP : INT := 50;
      c_NUM_ALARMS : INT := 15;
      c_AOI_MAX_RETRY : INT := 2;  (* Novas tentativas após a 1a falha *)
      c_AX_X : INT := 1;  (* Índices dos eixos *)
      c_AX_Y : INT := 2;
      c_AX_Z : INT := 3;
      c_AX_T : INT := 4;
      c_ALM_ESTOP : INT := 1;  (* Índices dos alarmes *)
      c_ALM_DOOR : INT := 2;
      c_ALM_HMI : INT := 3;
      c_ALM_CONVEYOR : INT := 4;
      c_ALM_AXIS_X : INT := 5;
      c_ALM_AXIS_Y : INT := 6;
      c_ALM_AXIS_Z : INT := 7;
      c_ALM_AXIS_T : INT := 8;
      c_ALM_CLAMP : INT := 9;
      c_ALM_STOPPER : INT := 10;
      c_ALM_PICK_FAIL : INT := 11;
      c_ALM_VAC_LOSS : INT := 12;
      c_ALM_AOI_TIMEOUT : INT := 13;
      c_ALM_RECIPE : INT := 14;
      c_ALM_Z_INTERLOCK : INT := 15;
      xEStopOk : BOOL;  (* TRUE = circuito de emergência íntegro (NF) *)
      xDoorClosed : BOOL;  (* TRUE = porta de proteção fechada (NF) *)
      xSensZ1 : BOOL;  (* Presença de placa: zona de entrada *)
      xSensZ2 : BOOL;  (* Presença de placa: zona de montagem *)
      xSensZ3 : BOOL;  (* Presença de placa: zona de saída/AOI *)
      xClampExtended : BOOL;  (* Grampo da zona 2: fim de curso avançado *)
      xClampRetracted : BOOL;  (* Grampo da zona 2: fim de curso recuado *)
      xStopExtended : BOOL;  (* Batente da zona 3: fim de curso avançado *)
      xStopRetracted : BOOL;  (* Batente da zona 3: fim de curso recuado *)
      xVacuumOk : BOOL;  (* Pressostato de vácuo *)
      xAoiDone : BOOL;  (* AOI: resultado disponível *)
      xAoiPass : BOOL;  (* AOI: TRUE = aprovada *)
      xSmemaUpAvail : BOOL;  (* SMEMA a montante: placa disponível *)
      xSmemaDownReady : BOOL;  (* SMEMA a jusante: máquina pronta *)
      xAxisDriveReady : ARRAY[1..4] OF BOOL;
      xAxisDriveFault : ARRAY[1..4] OF BOOL;
      xAxisHomeDone : ARRAY[1..4] OF BOOL;
      rAxisActPos : ARRAY[1..4] OF REAL;  (* Posição real [mm | graus] *)
      xMotor1 : BOOL;  (* Motor esteira zona 1 *)
      xMotor2 : BOOL;  (* Motor esteira zona 2 *)
      xMotor3 : BOOL;  (* Motor esteira zona 3 *)
      xClampValve : BOOL;  (* Válvula do grampo (mola de retorno) *)
      xStopValve : BOOL;  (* Válvula do batente (mola de retorno) *)
      xVacValve : BOOL;  (* Vácuo do cabeçote *)
      xBlowValve : BOOL;  (* Sopro de liberação *)
      xAoiTrigger : BOOL;  (* Disparo da inspeção *)
      xSmemaUpReady : BOOL;  (* SMEMA a montante: máquina pronta *)
      xSmemaDownAvail : BOOL;  (* SMEMA a jusante: placa disponível *)
      xBoardRejectedOut : BOOL;  (* Placa em saída foi rejeitada *)
      xAxisPower : ARRAY[1..4] OF BOOL;
      xAxisHome : ARRAY[1..4] OF BOOL;
      xAxisExecute : ARRAY[1..4] OF BOOL;
      rAxisSetpoint : ARRAY[1..4] OF REAL;
      rAxisMin : ARRAY[1..4] OF REAL := [0.0, 0.0, 0.0, -180.0];
      rAxisMax : ARRAY[1..4] OF REAL := [300.0, 250.0, 50.0, 180.0];
      rZSafe : REAL := 40.0;  (* Altura segura para deslocamento XY *)
      rZPick : REAL := 5.0;  (* Altura de coleta *)
      rZPlace : REAL := 8.0;  (* Altura de montagem *)
      rZTol : REAL := 1.0;  (* Tolerância da altura segura *)
      rParkX : REAL := 0.0;  (* Posição de repouso *)
      rParkY : REAL := 0.0;
      rParkT : REAL := 0.0;
      tCylTimeout : TIME := TIME#2s0ms;  (* Tempo máximo de movimento dos cilindros *)
      tConvTimeout : TIME := TIME#15s0ms;  (* Tempo máximo de transferência de placa *)
      tVacConfirm : TIME := TIME#1s0ms;  (* Tempo máximo para confirmar a pega *)
      tHmiTimeout : TIME := TIME#3s0ms;  (* Tempo sem heartbeat da IHM *)
      tAoiTimeout : TIME := TIME#10s0ms;  (* Tempo máximo de resposta da AOI *)
      iHmiHeartbeat : UINT;  (* IHM incrementa/alterna periodicamente *)
      xCmdStart : BOOL;
      xCmdStop : BOOL;
      xCmdHome : BOOL;
      xCmdAck : BOOL;
      xCmdReset : BOOL;
      xCmdClearZones : BOOL;  (* Ressincroniza zonas pelos sensores (máquina parada) *)
      xCmdResetCounters : BOOL;
      xCmdRecipeSel : BOOL;  (* Borda de subida: seleciona receita *)
      iRecipeReq : INT;  (* Receita pedida (1..3) *)
      iRecipeActive : INT;
      xRecipeValid : BOOL;
      xRecipeRejected : BOOL;  (* Troca recusada: máquina em operação *)
      eMachineState : E_MachineState := E_MachineState.INIT;
      xAlarmActive : ARRAY[1..15] OF BOOL;
      xAlarmAcked : ARRAY[1..15] OF BOOL;
      xAnyAlarm : BOOL;
      xAnyUnacked : BOOL;
      xSafetyOk : BOOL;  (* Emergência e porta OK (com atraso de rearme) *)
      xHmiOk : BOOL;
      xDrivesEnable : BOOL;
      xAutoEnable : BOOL;  (* Ciclo automático liberado *)
      xMotionRun : BOOL;  (* Serviços de movimento liberados *)
      xResetPulse : BOOL;  (* Pulso de reset para os dispositivos *)
      xStartRefusedRecipe : BOOL;  (* Pulso: partida recusada, receita inválida *)
      xHomeReq : BOOL;  (* Serviços de movimento *)
      xHomeSeqDone : BOOL;
      xAllHomed : BOOL;
      xMoveXYTReq : BOOL;
      xXYTDone : BOOL;
      xMoveZReq : BOOL;
      xZDone : BOOL;
      rTgtX : REAL;
      rTgtY : REAL;
      rTgtZ : REAL;
      rTgtT : REAL;
      xAxisFault : ARRAY[1..4] OF BOOL;
      xMotionFault : BOOL;
      xZInterlockFault : BOOL;
      xBoardInAsm : BOOL;  (* Placa posicionada na zona de montagem *)
      xAsmDone : BOOL;  (* Montagem concluída: libera a placa *)
      xBoardInInsp : BOOL;  (* Placa posicionada na zona de inspeção *)
      xInspDone : BOOL;  (* Inspeção concluída: libera a placa *)
      xCurBoardRejected : BOOL;
      xConveyorFault : BOOL;
      xClampFault : BOOL;  (* Pneumática, vácuo e AOI *)
      xStopperFault : BOOL;
      xPickFail : BOOL;
      xGripLoss : BOOL;
      xAoiTimeout : BOOL;
      aRecipes : ARRAY[1..3] OF ST_Recipe;
      diBoardsProduced : DINT;  (* Placas que concluíram o ciclo (aprovadas + rejeitadas) *)
      diBoardsRejected : DINT;  (* Placas rejeitadas (subconjunto das produzidas) *)
    END_VAR
    TASK MainTask(INTERVAL := T#20ms, PRIORITY := 1);
    PROGRAM PRG_Safety WITH MainTask : PRG_Safety;
    PROGRAM PRG_Motion WITH MainTask : PRG_Motion;
    PROGRAM PRG_PickPlace WITH MainTask : PRG_PickPlace;
    PROGRAM PRG_Main WITH MainTask : PRG_Main;
    PROGRAM PRG_Conveyor WITH MainTask : PRG_Conveyor;
    PROGRAM PRG_AOI WITH MainTask : PRG_AOI;
    PROGRAM PRG_Alarms WITH MainTask : PRG_Alarms;
  END_RESOURCE
END_CONFIGURATION
